Fanuc TP program (LS listing): Dispensing.LS

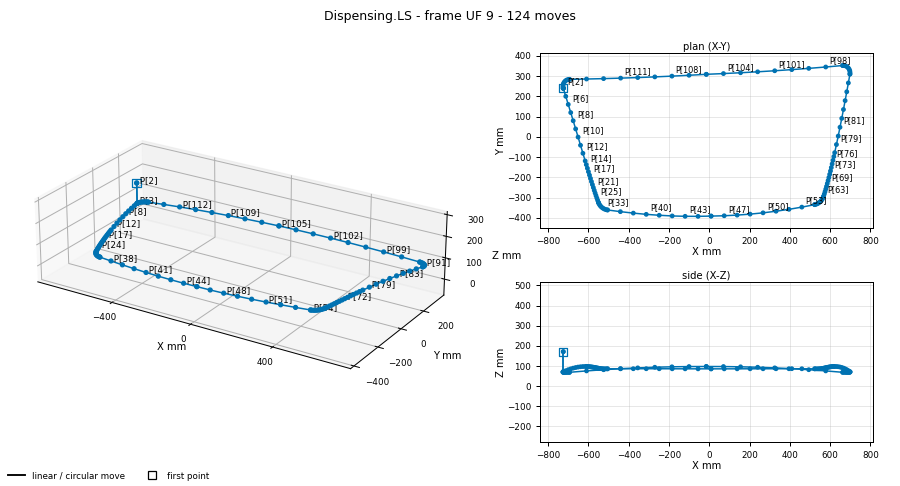
[picture p0: tool path of Dispensing.LS in frame UF 9, 124 of 125 moves have a stored position in this frame; points joined in program order, loops and branches not executed]
/PROG  Dispensing
/ATTR
OWNER		= MNEDITOR;
COMMENT		= "RoboDK sequence";
PROG_SIZE	= 0;
CREATE		= DATE 31-12-14  TIME 12:00:00;
MODIFIED	= DATE 31-12-14  TIME 12:00:00;
FILE_NAME	= Dispensing;
VERSION		= 0;
LINE_COUNT	= 145;
MEMORY_SIZE	= 0;
PROTECT		= READ_WRITE;
TCD:  STACK_SIZE	= 0,
      TASK_PRIORITY	= 50,
      TIME_SLICE	= 0,
      BUSY_LAMP_OFF	= 0,
      ABORT_REQUEST	= 0,
      PAUSE_REQUEST	= 0;
DEFAULT_GROUP	= 1,*,*,*,*,*,*;
CONTROL_CODE	= 00000000 00000000;
/MN
   1:  ! Program generated by VerticalBot Studio for Fanuc M-710iC/45M ;
   2:  ! on 25/10/2026 12:00:00 ;
   3:  ! Using nominal kinematics. ;
   4:  PR[9,1]=1.091 ;
   5:  PR[9,2]=1290.750 ;
   6:  PR[9,3]=1139.170 ;
   7:  PR[9,4]=-158.040 ;
   8:  PR[9,5]=0.000 ;
   9:  PR[9,6]=-180.000 ;
  10:  UFRAME[9]=PR[9] ;
  11:  UFRAME_NUM=9 ;
  12:  PR[9,1]=0.000 ;
  13:  PR[9,2]=0.000 ;
  14:  PR[9,3]=0.000 ;
  15:  PR[9,4]=0.000 ;
  16:  PR[9,5]=0.000 ;
  17:  PR[9,6]=0.000 ;
  18:  UTOOL[9]=PR[9] ;
  19:  UTOOL_NUM=9 ;
  20:  ! show Car windshield ;
  21:J P[1] 20% FINE ;
  22:L P[2] 1000mm/sec FINE ;
  23:L P[3] 1000mm/sec FINE ;
  24:L P[4] 1000mm/sec FINE ;
  25:L P[5] 50mm/sec FINE ;
  26:L P[6] 50mm/sec FINE ;
  27:L P[7] 50mm/sec FINE ;
  28:L P[8] 50mm/sec FINE ;
  29:L P[9] 50mm/sec FINE ;
  30:L P[10] 50mm/sec FINE ;
  31:L P[11] 50mm/sec FINE ;
  32:L P[12] 50mm/sec FINE ;
  33:L P[13] 50mm/sec FINE ;
  34:L P[14] 50mm/sec FINE ;
  35:L P[15] 50mm/sec FINE ;
  36:L P[16] 50mm/sec FINE ;
  37:L P[17] 50mm/sec FINE ;
  38:L P[18] 50mm/sec FINE ;
  39:L P[19] 50mm/sec FINE ;
  40:L P[20] 50mm/sec FINE ;
  41:L P[21] 50mm/sec FINE ;
  42:L P[22] 50mm/sec FINE ;
  43:L P[23] 50mm/sec FINE ;
  44:L P[24] 50mm/sec FINE ;
  45:L P[25] 50mm/sec FINE ;
  46:L P[26] 50mm/sec FINE ;
  47:L P[27] 50mm/sec FINE ;
  48:L P[28] 50mm/sec FINE ;
  49:L P[29] 50mm/sec FINE ;
  50:L P[30] 50mm/sec FINE ;
  51:L P[31] 50mm/sec FINE ;
  52:L P[32] 50mm/sec FINE ;
  53:L P[33] 50mm/sec FINE ;
  54:L P[34] 50mm/sec FINE ;
  55:L P[35] 50mm/sec FINE ;
  56:L P[36] 50mm/sec FINE ;
  57:L P[37] 50mm/sec FINE ;
  58:L P[38] 50mm/sec FINE ;
  59:L P[39] 50mm/sec FINE ;
  60:L P[40] 50mm/sec FINE ;
  61:L P[41] 50mm/sec FINE ;
  62:L P[42] 50mm/sec FINE ;
  63:L P[43] 50mm/sec FINE ;
  64:L P[44] 50mm/sec FINE ;
  65:L P[45] 50mm/sec FINE ;
  66:L P[46] 50mm/sec FINE ;
  67:L P[47] 50mm/sec FINE ;
  68:L P[48] 50mm/sec FINE ;
  69:L P[49] 50mm/sec FINE ;
  70:L P[50] 50mm/sec FINE ;
  71:L P[51] 50mm/sec FINE ;
  72:L P[52] 50mm/sec FINE ;
  73:L P[53] 50mm/sec FINE ;
  74:L P[54] 50mm/sec FINE ;
  75:L P[55] 50mm/sec FINE ;
  76:L P[56] 50mm/sec FINE ;
  77:L P[57] 50mm/sec FINE ;
  78:L P[58] 50mm/sec FINE ;
  79:L P[59] 50mm/sec FINE ;
  80:L P[60] 50mm/sec FINE ;
  81:L P[61] 50mm/sec FINE ;
  82:L P[62] 50mm/sec FINE ;
  83:L P[63] 50mm/sec FINE ;
  84:L P[64] 50mm/sec FINE ;
  85:L P[65] 50mm/sec FINE ;
  86:L P[66] 50mm/sec FINE ;
  87:L P[67] 50mm/sec FINE ;
  88:L P[68] 50mm/sec FINE ;
  89:L P[69] 50mm/sec FINE ;
  90:L P[70] 50mm/sec FINE ;
  91:L P[71] 50mm/sec FINE ;
  92:L P[72] 50mm/sec FINE ;
  93:L P[73] 50mm/sec FINE ;
  94:L P[74] 50mm/sec FINE ;
  95:L P[75] 50mm/sec FINE ;
  96:L P[76] 50mm/sec FINE ;
  97:L P[77] 50mm/sec FINE ;
  98:L P[78] 50mm/sec FINE ;
  99:L P[79] 50mm/sec FINE ;
 100:L P[80] 50mm/sec FINE ;
 101:L P[81] 50mm/sec FINE ;
 102:L P[82] 50mm/sec FINE ;
 103:L P[83] 50mm/sec FINE ;
 104:L P[84] 50mm/sec FINE ;
 105:L P[85] 50mm/sec FINE ;
 106:L P[86] 50mm/sec FINE ;
 107:L P[87] 50mm/sec FINE ;
 108:L P[88] 50mm/sec FINE ;
 109:L P[89] 50mm/sec FINE ;
 110:L P[90] 50mm/sec FINE ;
 111:L P[91] 50mm/sec FINE ;
 112:L P[92] 50mm/sec FINE ;
 113:L P[93] 50mm/sec FINE ;
 114:L P[94] 50mm/sec FINE ;
 115:L P[95] 50mm/sec FINE ;
 116:L P[96] 50mm/sec FINE ;
 117:L P[97] 50mm/sec FINE ;
 118:L P[98] 50mm/sec FINE ;
 119:L P[99] 50mm/sec FINE ;
 120:L P[100] 50mm/sec FINE ;
 121:L P[101] 50mm/sec FINE ;
 122:L P[102] 50mm/sec FINE ;
 123:L P[103] 50mm/sec FINE ;
 124:L P[104] 50mm/sec FINE ;
 125:L P[105] 50mm/sec FINE ;
 126:L P[106] 50mm/sec FINE ;
 127:L P[107] 50mm/sec FINE ;
 128:L P[108] 50mm/sec FINE ;
 129:L P[109] 50mm/sec FINE ;
 130:L P[110] 50mm/sec FINE ;
 131:L P[111] 50mm/sec FINE ;
 132:L P[112] 50mm/sec FINE ;
 133:L P[113] 50mm/sec FINE ;
 134:L P[114] 50mm/sec FINE ;
 135:L P[115] 50mm/sec FINE ;
 136:L P[116] 50mm/sec FINE ;
 137:L P[117] 50mm/sec FINE ;
 138:L P[118] 50mm/sec FINE ;
 139:L P[119] 50mm/sec FINE ;
 140:L P[120] 50mm/sec FINE ;
 141:L P[121] 50mm/sec FINE ;
 142:L P[122] 50mm/sec FINE ;
 143:L P[123] 50mm/sec FINE ;
 144:L P[124] 1000mm/sec FINE ;
 145:L P[125] 1000mm/sec FINE ;
/POS
P[1]{
   GP1:
    UF : 9, UT : 9,
	J1=    62.093 deg,	J2=    9.692 deg,	J3=    -25.783 deg,
	J4=    -167.561 deg,	J5=    -102.814 deg,	J6=    -22.106 deg
};
P[2]{
   GP1:
    UF : 9, UT : 9,        CONFIG : 'F U T, 0, 0, 0',
	X =  -725.181  mm,	Y =   240.604  mm,	Z =   171.303  mm,
	W =   175.329 deg,	P =     5.366 deg,	R =    92.372 deg
};
P[3]{
   GP1:
    UF : 9, UT : 9,        CONFIG : 'F U T, 0, 0, 0',
	X =  -725.181  mm,	Y =   240.604  mm,	Z =    71.303  mm,
	W =   175.329 deg,	P =     5.366 deg,	R =    92.372 deg
};
P[4]{
   GP1:
    UF : 9, UT : 9,        CONFIG : 'F U T, 0, 0, 0',
	X =  -725.181  mm,	Y =   240.604  mm,	Z =    71.303  mm,
	W =   175.329 deg,	P =     5.366 deg,	R =    92.372 deg
};
P[5]{
   GP1:
    UF : 9, UT : 9,        CONFIG : 'F U T, 0, 0, 0',
	X =  -712.750  mm,	Y =   200.498  mm,	Z =    76.770  mm,
	W =   175.467 deg,	P =     4.506 deg,	R =    92.372 deg
};
P[6]{
   GP1:
    UF : 9, UT : 9,        CONFIG : 'F U T, 0, 0, 0',
	X =  -700.389  mm,	Y =   160.323  mm,	Z =    81.631  mm,
	W =   175.606 deg,	P =     3.637 deg,	R =    92.368 deg
};
P[7]{
   GP1:
    UF : 9, UT : 9,        CONFIG : 'F U T, 0, 0, 0',
	X =  -688.092  mm,	Y =   120.075  mm,	Z =    85.874  mm,
	W =   175.745 deg,	P =     2.761 deg,	R =    92.358 deg
};
P[8]{
   GP1:
    UF : 9, UT : 9,        CONFIG : 'F U T, 0, 0, 0',
	X =  -675.855  mm,	Y =    79.754  mm,	Z =    89.484  mm,
	W =   175.884 deg,	P =     1.877 deg,	R =    92.344 deg
};
P[9]{
   GP1:
    UF : 9, UT : 9,        CONFIG : 'F U T, 0, 0, 0',
	X =  -663.685  mm,	Y =    39.408  mm,	Z =    92.446  mm,
	W =   176.023 deg,	P =     0.988 deg,	R =    92.324 deg
};
P[10]{
   GP1:
    UF : 9, UT : 9,        CONFIG : 'F U T, 0, 0, 0',
	X =  -651.566  mm,	Y =    -0.954  mm,	Z =    94.751  mm,
	W =   176.161 deg,	P =     0.093 deg,	R =    92.300 deg
};
P[11]{
   GP1:
    UF : 9, UT : 9,        CONFIG : 'F U T, 0, 0, 0',
	X =  -639.480  mm,	Y =   -41.336  mm,	Z =    96.391  mm,
	W =   176.300 deg,	P =    -0.807 deg,	R =    92.270 deg
};
P[12]{
   GP1:
    UF : 9, UT : 9,        CONFIG : 'F U T, 0, 0, 0',
	X =  -627.611  mm,	Y =   -81.041  mm,	Z =    97.348  mm,
	W =   176.437 deg,	P =    -1.696 deg,	R =    92.236 deg
};
P[13]{
   GP1:
    UF : 9, UT : 9,        CONFIG : 'F U T, 0, 0, 0',
	X =  -616.257  mm,	Y =  -118.952  mm,	Z =    97.652  mm,
	W =   176.568 deg,	P =    -2.548 deg,	R =    92.199 deg
};
P[14]{
   GP1:
    UF : 9, UT : 9,        CONFIG : 'F U T, 0, 0, 0',
	X =  -610.772  mm,	Y =  -137.196  mm,	Z =    97.583  mm,
	W =   176.632 deg,	P =    -2.960 deg,	R =    92.180 deg
};
P[15]{
   GP1:
    UF : 9, UT : 9,        CONFIG : 'F U T, 0, 0, 0',
	X =  -605.414  mm,	Y =  -154.948  mm,	Z =    97.382  mm,
	W =   176.693 deg,	P =    -3.361 deg,	R =    92.160 deg
};
P[16]{
   GP1:
    UF : 9, UT : 9,        CONFIG : 'F U T, 0, 0, 0',
	X =  -600.181  mm,	Y =  -172.192  mm,	Z =    97.059  mm,
	W =   176.753 deg,	P =    -3.751 deg,	R =    92.140 deg
};
P[17]{
   GP1:
    UF : 9, UT : 9,        CONFIG : 'F U T, 0, 0, 0',
	X =  -595.071  mm,	Y =  -188.915  mm,	Z =    96.626  mm,
	W =   176.812 deg,	P =    -4.130 deg,	R =    92.119 deg
};
P[18]{
   GP1:
    UF : 9, UT : 9,        CONFIG : 'F U T, 0, 0, 0',
	X =  -590.085  mm,	Y =  -205.104  mm,	Z =    96.094  mm,
	W =   176.869 deg,	P =    -4.497 deg,	R =    92.098 deg
};
P[19]{
   GP1:
    UF : 9, UT : 9,        CONFIG : 'F U T, 0, 0, 0',
	X =  -585.219  mm,	Y =  -220.743  mm,	Z =    95.475  mm,
	W =   176.924 deg,	P =    -4.853 deg,	R =    92.077 deg
};
P[20]{
   GP1:
    UF : 9, UT : 9,        CONFIG : 'F U T, 0, 0, 0',
	X =  -580.473  mm,	Y =  -235.820  mm,	Z =    94.782  mm,
	W =   176.977 deg,	P =    -5.196 deg,	R =    92.056 deg
};
P[21]{
   GP1:
    UF : 9, UT : 9,        CONFIG : 'F U T, 0, 0, 0',
	X =  -575.845  mm,	Y =  -250.320  mm,	Z =    94.024  mm,
	W =   177.029 deg,	P =    -5.527 deg,	R =    92.035 deg
};
P[22]{
   GP1:
    UF : 9, UT : 9,        CONFIG : 'F U T, 0, 0, 0',
	X =  -571.333  mm,	Y =  -264.228  mm,	Z =    93.215  mm,
	W =   177.079 deg,	P =    -5.844 deg,	R =    92.015 deg
};
P[23]{
   GP1:
    UF : 9, UT : 9,        CONFIG : 'F U T, 0, 0, 0',
	X =  -566.936  mm,	Y =  -277.532  mm,	Z =    92.366  mm,
	W =   177.127 deg,	P =    -6.149 deg,	R =    91.994 deg
};
P[24]{
   GP1:
    UF : 9, UT : 9,        CONFIG : 'F U T, 0, 0, 0',
	X =  -562.651  mm,	Y =  -290.217  mm,	Z =    91.488  mm,
	W =   177.173 deg,	P =    -6.439 deg,	R =    91.974 deg
};
P[25]{
   GP1:
    UF : 9, UT : 9,        CONFIG : 'F U T, 0, 0, 0',
	X =  -558.477  mm,	Y =  -302.269  mm,	Z =    90.592  mm,
	W =   177.217 deg,	P =    -6.715 deg,	R =    91.954 deg
};
P[26]{
   GP1:
    UF : 9, UT : 9,        CONFIG : 'F U T, 0, 0, 0',
	X =  -554.411  mm,	Y =  -313.674  mm,	Z =    89.688  mm,
	W =   177.260 deg,	P =    -6.977 deg,	R =    91.935 deg
};
P[27]{
   GP1:
    UF : 9, UT : 9,        CONFIG : 'F U T, 0, 0, 0',
	X =  -550.453  mm,	Y =  -324.419  mm,	Z =    88.788  mm,
	W =   177.300 deg,	P =    -7.225 deg,	R =    91.917 deg
};
P[28]{
   GP1:
    UF : 9, UT : 9,        CONFIG : 'F U T, 0, 0, 0',
	X =  -550.453  mm,	Y =  -324.419  mm,	Z =    88.788  mm,
	W =   177.300 deg,	P =    -7.225 deg,	R =    91.917 deg
};
P[29]{
   GP1:
    UF : 9, UT : 9,        CONFIG : 'F U T, 0, 0, 0',
	X =  -547.304  mm,	Y =  -331.418  mm,	Z =    88.190  mm,
	W =   177.329 deg,	P =    -7.387 deg,	R =    91.904 deg
};
P[30]{
   GP1:
    UF : 9, UT : 9,        CONFIG : 'F U T, 0, 0, 0',
	X =  -543.300  mm,	Y =  -337.927  mm,	Z =    87.644  mm,
	W =   177.361 deg,	P =    -7.542 deg,	R =    91.891 deg
};
P[31]{
   GP1:
    UF : 9, UT : 9,        CONFIG : 'F U T, 0, 0, 0',
	X =  -538.489  mm,	Y =  -343.856  mm,	Z =    87.159  mm,
	W =   177.396 deg,	P =    -7.686 deg,	R =    91.879 deg
};
P[32]{
   GP1:
    UF : 9, UT : 9,        CONFIG : 'F U T, 0, 0, 0',
	X =  -532.947  mm,	Y =  -349.088  mm,	Z =    86.749  mm,
	W =   177.432 deg,	P =    -7.817 deg,	R =    91.866 deg
};
P[33]{
   GP1:
    UF : 9, UT : 9,        CONFIG : 'F U T, 0, 0, 0',
	X =  -526.769  mm,	Y =  -353.519  mm,	Z =    86.427  mm,
	W =   177.469 deg,	P =    -7.932 deg,	R =    91.855 deg
};
P[34]{
   GP1:
    UF : 9, UT : 9,        CONFIG : 'F U T, 0, 0, 0',
	X =  -520.043  mm,	Y =  -357.070  mm,	Z =    86.201  mm,
	W =   177.506 deg,	P =    -8.029 deg,	R =    91.844 deg
};
P[35]{
   GP1:
    UF : 9, UT : 9,        CONFIG : 'F U T, 0, 0, 0',
	X =  -512.920  mm,	Y =  -359.651  mm,	Z =    86.084  mm,
	W =   177.544 deg,	P =    -8.106 deg,	R =    91.834 deg
};
P[36]{
   GP1:
    UF : 9, UT : 9,        CONFIG : 'F U T, 0, 0, 0',
	X =  -505.502  mm,	Y =  -361.220  mm,	Z =    86.081  mm,
	W =   177.580 deg,	P =    -8.161 deg,	R =    91.826 deg
};
P[37]{
   GP1:
    UF : 9, UT : 9,        CONFIG : 'F U T, 0, 0, 0',
	X =  -505.502  mm,	Y =  -361.220  mm,	Z =    86.081  mm,
	W =   177.580 deg,	P =    -8.161 deg,	R =    91.826 deg
};
P[38]{
   GP1:
    UF : 9, UT : 9,        CONFIG : 'F U T, 0, 0, 0',
	X =  -441.508  mm,	Y =  -369.591  mm,	Z =    86.422  mm,
	W =   177.879 deg,	P =    -8.515 deg,	R =    91.761 deg
};
P[39]{
   GP1:
    UF : 9, UT : 9,        CONFIG : 'F U T, 0, 0, 0',
	X =  -377.427  mm,	Y =  -376.823  mm,	Z =    86.546  mm,
	W =   178.169 deg,	P =    -8.829 deg,	R =    91.696 deg
};
P[40]{
   GP1:
    UF : 9, UT : 9,        CONFIG : 'F U T, 0, 0, 0',
	X =  -313.197  mm,	Y =  -382.829  mm,	Z =    86.519  mm,
	W =   178.450 deg,	P =    -9.101 deg,	R =    91.633 deg
};
P[41]{
   GP1:
    UF : 9, UT : 9,        CONFIG : 'F U T, 0, 0, 0',
	X =  -248.757  mm,	Y =  -387.517  mm,	Z =    86.400  mm,
	W =   178.724 deg,	P =    -9.328 deg,	R =    91.572 deg
};
P[42]{
   GP1:
    UF : 9, UT : 9,        CONFIG : 'F U T, 0, 0, 0',
	X =  -184.353  mm,	Y =  -390.786  mm,	Z =    86.237  mm,
	W =   178.990 deg,	P =    -9.507 deg,	R =    91.514 deg
};
P[43]{
   GP1:
    UF : 9, UT : 9,        CONFIG : 'F U T, 0, 0, 0',
	X =  -120.125  mm,	Y =  -392.569  mm,	Z =    86.084  mm,
	W =   179.250 deg,	P =    -9.637 deg,	R =    91.460 deg
};
P[44]{
   GP1:
    UF : 9, UT : 9,        CONFIG : 'F U T, 0, 0, 0',
	X =   -55.881  mm,	Y =  -392.821  mm,	Z =    85.977  mm,
	W =   179.506 deg,	P =    -9.716 deg,	R =    91.410 deg
};
P[45]{
   GP1:
    UF : 9, UT : 9,        CONFIG : 'F U T, 0, -1, 0',
	X =     8.571  mm,	Y =  -391.495  mm,	Z =    85.934  mm,
	W =   179.760 deg,	P =    -9.744 deg,	R =    91.365 deg
};
P[46]{
   GP1:
    UF : 9, UT : 9,        CONFIG : 'F U T, 0, -1, 0',
	X =     9.058  mm,	Y =  -391.485  mm,	Z =    85.935  mm,
	W =  -180.000 deg,	P =    -9.745 deg,	R =    91.325 deg
};
P[47]{
   GP1:
    UF : 9, UT : 9,        CONFIG : 'F U T, 0, -1, 0',
	X =    73.885  mm,	Y =  -389.871  mm,	Z =    85.968  mm,
	W =  -179.506 deg,	P =    -9.718 deg,	R =    91.246 deg
};
P[48]{
   GP1:
    UF : 9, UT : 9,        CONFIG : 'F U T, 0, -1, 0',
	X =   138.144  mm,	Y =  -386.662  mm,	Z =    86.067  mm,
	W =  -179.251 deg,	P =    -9.640 deg,	R =    91.212 deg
};
P[49]{
   GP1:
    UF : 9, UT : 9,        CONFIG : 'F U T, 0, -1, 0',
	X =   202.382  mm,	Y =  -381.853  mm,	Z =    86.213  mm,
	W =  -178.991 deg,	P =    -9.511 deg,	R =    91.185 deg
};
P[50]{
   GP1:
    UF : 9, UT : 9,        CONFIG : 'F U T, 0, -1, 0',
	X =   266.788  mm,	Y =  -375.443  mm,	Z =    86.368  mm,
	W =  -178.725 deg,	P =    -9.333 deg,	R =    91.164 deg
};
P[51]{
   GP1:
    UF : 9, UT : 9,        CONFIG : 'F U T, 0, -1, 0',
	X =   331.224  mm,	Y =  -367.474  mm,	Z =    86.482  mm,
	W =  -178.451 deg,	P =    -9.107 deg,	R =    91.149 deg
};
P[52]{
   GP1:
    UF : 9, UT : 9,        CONFIG : 'F U T, 0, -1, 0',
	X =   395.430  mm,	Y =  -358.032  mm,	Z =    86.504  mm,
	W =  -178.170 deg,	P =    -8.837 deg,	R =    91.142 deg
};
P[53]{
   GP1:
    UF : 9, UT : 9,        CONFIG : 'F U T, 0, -1, 0',
	X =   459.460  mm,	Y =  -347.178  mm,	Z =    86.377  mm,
	W =  -177.881 deg,	P =    -8.524 deg,	R =    91.142 deg
};
P[54]{
   GP1:
    UF : 9, UT : 9,        CONFIG : 'F U T, 0, -1, 0',
	X =   523.365  mm,	Y =  -334.972  mm,	Z =    86.033  mm,
	W =  -177.582 deg,	P =    -8.171 deg,	R =    91.150 deg
};
P[55]{
   GP1:
    UF : 9, UT : 9,        CONFIG : 'F U T, 0, -1, 0',
	X =   523.365  mm,	Y =  -334.972  mm,	Z =    86.033  mm,
	W =  -177.582 deg,	P =    -8.171 deg,	R =    91.150 deg
};
P[56]{
   GP1:
    UF : 9, UT : 9,        CONFIG : 'F U T, 0, -1, 0',
	X =   530.760  mm,	Y =  -332.922  mm,	Z =    86.036  mm,
	W =  -177.546 deg,	P =    -8.116 deg,	R =    91.153 deg
};
P[57]{
   GP1:
    UF : 9, UT : 9,        CONFIG : 'F U T, 0, -1, 0',
	X =   537.824  mm,	Y =  -329.835  mm,	Z =    86.153  mm,
	W =  -177.508 deg,	P =    -8.040 deg,	R =    91.159 deg
};
P[58]{
   GP1:
    UF : 9, UT : 9,        CONFIG : 'F U T, 0, -1, 0',
	X =   544.463  mm,	Y =  -325.760  mm,	Z =    86.379  mm,
	W =  -177.471 deg,	P =    -7.943 deg,	R =    91.168 deg
};
P[59]{
   GP1:
    UF : 9, UT : 9,        CONFIG : 'F U T, 0, -1, 0',
	X =   550.537  mm,	Y =  -320.790  mm,	Z =    86.702  mm,
	W =  -177.434 deg,	P =    -7.828 deg,	R =    91.180 deg
};
P[60]{
   GP1:
    UF : 9, UT : 9,        CONFIG : 'F U T, 0, -1, 0',
	X =   555.942  mm,	Y =  -315.021  mm,	Z =    87.112  mm,
	W =  -177.398 deg,	P =    -7.698 deg,	R =    91.194 deg
};
P[61]{
   GP1:
    UF : 9, UT : 9,        CONFIG : 'F U T, 0, -1, 0',
	X =   560.600  mm,	Y =  -308.550  mm,	Z =    87.598  mm,
	W =  -177.363 deg,	P =    -7.554 deg,	R =    91.211 deg
};
P[62]{
   GP1:
    UF : 9, UT : 9,        CONFIG : 'F U T, 0, -1, 0',
	X =   564.423  mm,	Y =  -301.516  mm,	Z =    88.146  mm,
	W =  -177.331 deg,	P =    -7.399 deg,	R =    91.230 deg
};
P[63]{
   GP1:
    UF : 9, UT : 9,        CONFIG : 'F U T, 0, -1, 0',
	X =   567.363  mm,	Y =  -294.023  mm,	Z =    88.745  mm,
	W =  -177.302 deg,	P =    -7.236 deg,	R =    91.251 deg
};
P[64]{
   GP1:
    UF : 9, UT : 9,        CONFIG : 'F U T, 0, -1, 0',
	X =   567.363  mm,	Y =  -294.023  mm,	Z =    88.745  mm,
	W =  -177.302 deg,	P =    -7.236 deg,	R =    91.251 deg
};
P[65]{
   GP1:
    UF : 9, UT : 9,        CONFIG : 'F U T, 0, -1, 0',
	X =   570.932  mm,	Y =  -282.728  mm,	Z =    89.636  mm,
	W =  -177.262 deg,	P =    -6.992 deg,	R =    91.283 deg
};
P[66]{
   GP1:
    UF : 9, UT : 9,        CONFIG : 'F U T, 0, -1, 0',
	X =   574.565  mm,	Y =  -270.743  mm,	Z =    90.529  mm,
	W =  -177.220 deg,	P =    -6.734 deg,	R =    91.317 deg
};
P[67]{
   GP1:
    UF : 9, UT : 9,        CONFIG : 'F U T, 0, -1, 0',
	X =   578.260  mm,	Y =  -258.082  mm,	Z =    91.417  mm,
	W =  -177.177 deg,	P =    -6.461 deg,	R =    91.353 deg
};
P[68]{
   GP1:
    UF : 9, UT : 9,        CONFIG : 'F U T, 0, -1, 0',
	X =   582.016  mm,	Y =  -244.758  mm,	Z =    92.287  mm,
	W =  -177.131 deg,	P =    -6.175 deg,	R =    91.392 deg
};
P[69]{
   GP1:
    UF : 9, UT : 9,        CONFIG : 'F U T, 0, -1, 0',
	X =   585.831  mm,	Y =  -230.784  mm,	Z =    93.131  mm,
	W =  -177.083 deg,	P =    -5.875 deg,	R =    91.433 deg
};
P[70]{
   GP1:
    UF : 9, UT : 9,        CONFIG : 'F U T, 0, -1, 0',
	X =   589.704  mm,	Y =  -216.173  mm,	Z =    93.936  mm,
	W =  -177.034 deg,	P =    -5.562 deg,	R =    91.476 deg
};
P[71]{
   GP1:
    UF : 9, UT : 9,        CONFIG : 'F U T, 0, -1, 0',
	X =   593.633  mm,	Y =  -200.937  mm,	Z =    94.693  mm,
	W =  -176.983 deg,	P =    -5.236 deg,	R =    91.522 deg
};
P[72]{
   GP1:
    UF : 9, UT : 9,        CONFIG : 'F U T, 0, -1, 0',
	X =   597.616  mm,	Y =  -185.092  mm,	Z =    95.388  mm,
	W =  -176.930 deg,	P =    -4.897 deg,	R =    91.570 deg
};
P[73]{
   GP1:
    UF : 9, UT : 9,        CONFIG : 'F U T, 0, -1, 0',
	X =   601.651  mm,	Y =  -168.648  mm,	Z =    96.011  mm,
	W =  -176.876 deg,	P =    -4.547 deg,	R =    91.620 deg
};
P[74]{
   GP1:
    UF : 9, UT : 9,        CONFIG : 'F U T, 0, -1, 0',
	X =   605.737  mm,	Y =  -151.621  mm,	Z =    96.551  mm,
	W =  -176.820 deg,	P =    -4.184 deg,	R =    91.672 deg
};
P[75]{
   GP1:
    UF : 9, UT : 9,        CONFIG : 'F U T, 0, -1, 0',
	X =   609.871  mm,	Y =  -134.022  mm,	Z =    96.996  mm,
	W =  -176.762 deg,	P =    -3.810 deg,	R =    91.728 deg
};
P[76]{
   GP1:
    UF : 9, UT : 9,        CONFIG : 'F U T, 0, -1, 0',
	X =   614.051  mm,	Y =  -115.865  mm,	Z =    97.334  mm,
	W =  -176.703 deg,	P =    -3.425 deg,	R =    91.785 deg
};
P[77]{
   GP1:
    UF : 9, UT : 9,        CONFIG : 'F U T, 0, -1, 0',
	X =   618.276  mm,	Y =   -97.163  mm,	Z =    97.554  mm,
	W =  -176.642 deg,	P =    -3.029 deg,	R =    91.845 deg
};
P[78]{
   GP1:
    UF : 9, UT : 9,        CONFIG : 'F U T, 0, -1, 0',
	X =   622.544  mm,	Y =   -77.931  mm,	Z =    97.645  mm,
	W =  -176.579 deg,	P =    -2.623 deg,	R =    91.907 deg
};
P[79]{
   GP1:
    UF : 9, UT : 9,        CONFIG : 'F U T, 0, -1, 0',
	X =   631.198  mm,	Y =   -37.925  mm,	Z =    97.399  mm,
	W =  -176.450 deg,	P =    -1.780 deg,	R =    92.038 deg
};
P[80]{
   GP1:
    UF : 9, UT : 9,        CONFIG : 'F U T, 0, -1, 0',
	X =   639.996  mm,	Y =     4.045  mm,	Z =    96.514  mm,
	W =  -176.314 deg,	P =    -0.901 deg,	R =    92.179 deg
};
P[81]{
   GP1:
    UF : 9, UT : 9,        CONFIG : 'F U T, 0, -1, 0',
	X =   648.878  mm,	Y =    47.647  mm,	Z =    94.924  mm,
	W =  -176.174 deg,	P =     0.007 deg,	R =    92.329 deg
};
P[82]{
   GP1:
    UF : 9, UT : 9,        CONFIG : 'F U T, 0, -1, 0',
	X =   657.573  mm,	Y =    91.479  mm,	Z =    92.644  mm,
	W =  -176.033 deg,	P =     0.915 deg,	R =    92.482 deg
};
P[83]{
   GP1:
    UF : 9, UT : 9,        CONFIG : 'F U T, 0, -1, 0',
	X =   666.058  mm,	Y =   135.316  mm,	Z =    89.688  mm,
	W =  -175.892 deg,	P =     1.817 deg,	R =    92.638 deg
};
P[84]{
   GP1:
    UF : 9, UT : 9,        CONFIG : 'F U T, 0, -1, 0',
	X =   674.353  mm,	Y =   179.152  mm,	Z =    86.066  mm,
	W =  -175.751 deg,	P =     2.713 deg,	R =    92.797 deg
};
P[85]{
   GP1:
    UF : 9, UT : 9,        CONFIG : 'F U T, 0, -1, 0',
	X =   682.468  mm,	Y =   222.942  mm,	Z =    81.793  mm,
	W =  -175.610 deg,	P =     3.601 deg,	R =    92.959 deg
};
P[86]{
   GP1:
    UF : 9, UT : 9,        CONFIG : 'F U T, 0, -1, 0',
	X =   690.411  mm,	Y =   266.680  mm,	Z =    76.885  mm,
	W =  -175.469 deg,	P =     4.482 deg,	R =    93.123 deg
};
P[87]{
   GP1:
    UF : 9, UT : 9,        CONFIG : 'F U T, 0, -1, 0',
	X =   698.195  mm,	Y =   310.369  mm,	Z =    71.355  mm,
	W =  -175.328 deg,	P =     5.354 deg,	R =    93.289 deg
};
P[88]{
   GP1:
    UF : 9, UT : 9,        CONFIG : 'F U T, 0, -1, 0',
	X =   698.195  mm,	Y =   310.369  mm,	Z =    71.355  mm,
	W =  -175.328 deg,	P =     5.354 deg,	R =    93.289 deg
};
P[89]{
   GP1:
    UF : 9, UT : 9,        CONFIG : 'F U T, 0, -1, 0',
	X =   698.725  mm,	Y =   318.498  mm,	Z =    70.329  mm,
	W =  -175.308 deg,	P =     5.515 deg,	R =    93.320 deg
};
P[90]{
   GP1:
    UF : 9, UT : 9,        CONFIG : 'F U T, 0, -1, 0',
	X =   697.484  mm,	Y =   326.580  mm,	Z =    69.430  mm,
	W =  -175.298 deg,	P =     5.674 deg,	R =    93.349 deg
};
P[91]{
   GP1:
    UF : 9, UT : 9,        CONFIG : 'F U T, 0, -1, 0',
	X =   694.546  mm,	Y =   334.166  mm,	Z =    68.709  mm,
	W =  -175.300 deg,	P =     5.823 deg,	R =    93.374 deg
};
P[92]{
   GP1:
    UF : 9, UT : 9,        CONFIG : 'F U T, 0, -1, 0',
	X =   690.052  mm,	Y =   340.884  mm,	Z =    68.206  mm,
	W =  -175.314 deg,	P =     5.953 deg,	R =    93.396 deg
};
P[93]{
   GP1:
    UF : 9, UT : 9,        CONFIG : 'F U T, 0, -1, 0',
	X =   684.250  mm,	Y =   346.352  mm,	Z =    67.955  mm,
	W =  -175.339 deg,	P =     6.058 deg,	R =    93.411 deg
};
P[94]{
   GP1:
    UF : 9, UT : 9,        CONFIG : 'F U T, 0, -1, 0',
	X =   677.435  mm,	Y =   350.280  mm,	Z =    67.974  mm,
	W =  -175.374 deg,	P =     6.133 deg,	R =    93.420 deg
};
P[95]{
   GP1:
    UF : 9, UT : 9,        CONFIG : 'F U T, 0, -1, 0',
	X =   669.973  mm,	Y =   352.443  mm,	Z =    68.267  mm,
	W =  -175.416 deg,	P =     6.173 deg,	R =    93.422 deg
};
P[96]{
   GP1:
    UF : 9, UT : 9,        CONFIG : 'F U T, 0, -1, 0',
	X =   662.283  mm,	Y =   352.715  mm,	Z =    68.820  mm,
	W =  -175.464 deg,	P =     6.176 deg,	R =    93.417 deg
};
P[97]{
   GP1:
    UF : 9, UT : 9,        CONFIG : 'F U T, 0, -1, 0',
	X =   662.283  mm,	Y =   352.715  mm,	Z =    68.820  mm,
	W =  -175.464 deg,	P =     6.176 deg,	R =    93.417 deg
};
P[98]{
   GP1:
    UF : 9, UT : 9,        CONFIG : 'F U T, 0, -1, 0',
	X =   578.111  mm,	Y =   345.429  mm,	Z =    75.733  mm,
	W =  -176.004 deg,	P =     6.008 deg,	R =    93.326 deg
};
P[99]{
   GP1:
    UF : 9, UT : 9,        CONFIG : 'F U T, 0, -1, 0',
	X =   493.807  mm,	Y =   338.691  mm,	Z =    81.683  mm,
	W =  -176.541 deg,	P =     5.864 deg,	R =    93.243 deg
};
P[100]{
   GP1:
    UF : 9, UT : 9,        CONFIG : 'F U T, 0, -1, 0',
	X =   409.361  mm,	Y =   332.492  mm,	Z =    86.682  mm,
	W =  -177.074 deg,	P =     5.744 deg,	R =    93.167 deg
};
P[101]{
   GP1:
    UF : 9, UT : 9,        CONFIG : 'F U T, 0, -1, 0',
	X =   324.760  mm,	Y =   326.826  mm,	Z =    90.739  mm,
	W =  -177.604 deg,	P =     5.648 deg,	R =    93.097 deg
};
P[102]{
   GP1:
    UF : 9, UT : 9,        CONFIG : 'F U T, 0, -1, 0',
	X =   240.009  mm,	Y =   321.685  mm,	Z =    93.861  mm,
	W =  -178.132 deg,	P =     5.578 deg,	R =    93.032 deg
};
P[103]{
   GP1:
    UF : 9, UT : 9,        CONFIG : 'F U T, 0, -1, 0',
	X =   155.150  mm,	Y =   317.057  mm,	Z =    96.051  mm,
	W =  -178.659 deg,	P =     5.535 deg,	R =    92.973 deg
};
P[104]{
   GP1:
    UF : 9, UT : 9,        CONFIG : 'F U T, 0, -1, 0',
	X =    70.232  mm,	Y =   312.934  mm,	Z =    97.314  mm,
	W =  -179.184 deg,	P =     5.519 deg,	R =    92.917 deg
};
P[105]{
   GP1:
    UF : 9, UT : 9,        CONFIG : 'F U T, 0, 0, 0',
	X =   -14.695  mm,	Y =   309.308  mm,	Z =    97.649  mm,
	W =  -179.709 deg,	P =     5.530 deg,	R =    92.865 deg
};
P[106]{
   GP1:
    UF : 9, UT : 9,        CONFIG : 'F U T, 0, 0, 0',
	X =   -15.315  mm,	Y =   309.276  mm,	Z =    97.650  mm,
	W =  -180.000 deg,	P =     5.530 deg,	R =    92.836 deg
};
P[107]{
   GP1:
    UF : 9, UT : 9,        CONFIG : 'F U T, 0, 0, 0',
	X =  -100.650  mm,	Y =   304.544  mm,	Z =    97.307  mm,
	W =   179.185 deg,	P =     5.520 deg,	R =    92.753 deg
};
P[108]{
   GP1:
    UF : 9, UT : 9,        CONFIG : 'F U T, 0, 0, 0',
	X =  -185.568  mm,	Y =   300.318  mm,	Z =    96.038  mm,
	W =   178.660 deg,	P =     5.538 deg,	R =    92.702 deg
};
P[109]{
   GP1:
    UF : 9, UT : 9,        CONFIG : 'F U T, 0, 0, 0',
	X =  -270.506  mm,	Y =   296.560  mm,	Z =    93.841  mm,
	W =   178.133 deg,	P =     5.583 deg,	R =    92.652 deg
};
P[110]{
   GP1:
    UF : 9, UT : 9,        CONFIG : 'F U T, 0, 0, 0',
	X =  -355.415  mm,	Y =   293.260  mm,	Z =    90.713  mm,
	W =   177.605 deg,	P =     5.654 deg,	R =    92.603 deg
};
P[111]{
   GP1:
    UF : 9, UT : 9,        CONFIG : 'F U T, 0, 0, 0',
	X =  -440.250  mm,	Y =   290.409  mm,	Z =    86.650  mm,
	W =   177.075 deg,	P =     5.751 deg,	R =    92.554 deg
};
P[112]{
   GP1:
    UF : 9, UT : 9,        CONFIG : 'F U T, 0, 0, 0',
	X =  -525.010  mm,	Y =   287.994  mm,	Z =    81.644  mm,
	W =   176.542 deg,	P =     5.873 deg,	R =    92.504 deg
};
P[113]{
   GP1:
    UF : 9, UT : 9,        CONFIG : 'F U T, 0, 0, 0',
	X =  -609.705  mm,	Y =   285.998  mm,	Z =    75.688  mm,
	W =   176.005 deg,	P =     6.019 deg,	R =    92.452 deg
};
P[114]{
   GP1:
    UF : 9, UT : 9,        CONFIG : 'F U T, 0, 0, 0',
	X =  -694.346  mm,	Y =   284.407  mm,	Z =    68.768  mm,
	W =   175.465 deg,	P =     6.187 deg,	R =    92.397 deg
};
P[115]{
   GP1:
    UF : 9, UT : 9,        CONFIG : 'F U T, 0, 0, 0',
	X =  -694.346  mm,	Y =   284.407  mm,	Z =    68.768  mm,
	W =   175.465 deg,	P =     6.187 deg,	R =    92.397 deg
};
P[116]{
   GP1:
    UF : 9, UT : 9,        CONFIG : 'F U T, 0, 0, 0',
	X =  -701.956  mm,	Y =   283.369  mm,	Z =    68.214  mm,
	W =   175.417 deg,	P =     6.185 deg,	R =    92.392 deg
};
P[117]{
   GP1:
    UF : 9, UT : 9,        CONFIG : 'F U T, 0, 0, 0',
	X =  -709.119  mm,	Y =   280.562  mm,	Z =    67.921  mm,
	W =   175.375 deg,	P =     6.145 deg,	R =    92.386 deg
};
P[118]{
   GP1:
    UF : 9, UT : 9,        CONFIG : 'F U T, 0, 0, 0',
	X =  -715.428  mm,	Y =   276.159  mm,	Z =    67.900  mm,
	W =   175.340 deg,	P =     6.071 deg,	R =    92.382 deg
};
P[119]{
   GP1:
    UF : 9, UT : 9,        CONFIG : 'F U T, 0, 0, 0',
	X =  -720.569  mm,	Y =   270.391  mm,	Z =    68.150  mm,
	W =   175.315 deg,	P =     5.966 deg,	R =    92.378 deg
};
P[120]{
   GP1:
    UF : 9, UT : 9,        CONFIG : 'F U T, 0, 0, 0',
	X =  -724.262  mm,	Y =   263.585  mm,	Z =    68.651  mm,
	W =   175.301 deg,	P =     5.836 deg,	R =    92.375 deg
};
P[121]{
   GP1:
    UF : 9, UT : 9,        CONFIG : 'F U T, 0, 0, 0',
	X =  -726.324  mm,	Y =   256.079  mm,	Z =    69.373  mm,
	W =   175.299 deg,	P =     5.687 deg,	R =    92.373 deg
};
P[122]{
   GP1:
    UF : 9, UT : 9,        CONFIG : 'F U T, 0, 0, 0',
	X =  -726.638  mm,	Y =   248.280  mm,	Z =    70.274  mm,
	W =   175.308 deg,	P =     5.528 deg,	R =    92.372 deg
};
P[123]{
   GP1:
    UF : 9, UT : 9,        CONFIG : 'F U T, 0, 0, 0',
	X =  -725.181  mm,	Y =   240.604  mm,	Z =    71.303  mm,
	W =   175.329 deg,	P =     5.366 deg,	R =    92.372 deg
};
P[124]{
   GP1:
    UF : 9, UT : 9,        CONFIG : 'F U T, 0, 0, 0',
	X =  -725.181  mm,	Y =   240.604  mm,	Z =    71.303  mm,
	W =   175.329 deg,	P =     5.366 deg,	R =    92.372 deg
};
P[125]{
   GP1:
    UF : 9, UT : 9,        CONFIG : 'F U T, 0, 0, 0',
	X =  -725.181  mm,	Y =   240.604  mm,	Z =   171.303  mm,
	W =   175.329 deg,	P =     5.366 deg,	R =    92.372 deg
};
/END
